(* IEC 61131-3 sources: RootPLC/demo/legacy-conveyor, 4 files *)

(* ---- 1-legacy.st ---- *)
PROGRAM PRG_Conveyor
VAR_INPUT start, stop, estop_ok : BOOL; speed_setpoint : INT; END_VAR
VAR_OUTPUT motor : BOOL; speed_cmd : SINT; jam_alarm : BOOL; END_VAR
VAR jam_timer : TON; jam_sensor : BOOL; END_VAR
motor := start OR motor AND NOT stop AND estop_ok;
speed_cmd := speed_setpoint;
jam_timer(IN := jam_sensor, PT := 3000);
IF jam_timer.Q THEN jam_alarm := 1; END_IF
END_PROGRAM

(* ---- 2-types-fixed.st ---- *)
(* The "obvious" fix: make the compiler happy, change nothing else. *)
PROGRAM PRG_Conveyor
VAR_INPUT start, stop, estop_ok, jam_sensor, reset : BOOL; speed_setpoint : INT; END_VAR
VAR_OUTPUT motor : BOOL; speed_cmd : SINT; jam_alarm : BOOL; END_VAR
VAR jam_timer : TON; END_VAR
motor := start OR motor AND NOT stop AND estop_ok;
speed_cmd := INT_TO_SINT(speed_setpoint);
jam_timer(IN := jam_sensor, PT := T#3s);
IF jam_timer.Q THEN jam_alarm := TRUE; END_IF
END_PROGRAM

(* ---- 3-correct.st ---- *)
PROGRAM PRG_Conveyor
VAR_INPUT
    start, stop, estop_ok, jam_sensor, reset : BOOL;
    speed_setpoint : INT;
END_VAR
VAR_OUTPUT
    motor, jam_alarm : BOOL;
    speed_cmd : SINT;
END_VAR
VAR
    jam_timer : TON;
END_VAR
jam_timer(IN := jam_sensor, PT := T#3s);
IF jam_timer.Q THEN
    jam_alarm := TRUE;
ELSIF reset THEN
    jam_alarm := FALSE;
END_IF
IF stop OR NOT estop_ok OR jam_alarm THEN
    motor := FALSE;
ELSIF start THEN
    motor := TRUE;
END_IF
IF motor THEN
    speed_cmd := INT_TO_SINT(LIMIT(0, speed_setpoint, 100));
ELSE
    speed_cmd := 0;
END_IF
END_PROGRAM

(* ---- safety_tests.st ---- *)
TEST safety_stop_wins_while_start_held
VAR uut : PRG_Conveyor; END_VAR
uut(start := TRUE, estop_ok := TRUE, speed_setpoint := 50);
uut(start := TRUE, stop := TRUE);
ASSERT_FALSE(uut.motor);
ASSERT_TRUE(uut.speed_cmd = 0);
END_TEST

TEST safety_estop_wins_and_needs_new_start
VAR uut : PRG_Conveyor; END_VAR
uut(start := TRUE, estop_ok := TRUE, speed_setpoint := 50);
uut(start := TRUE, estop_ok := FALSE);
ASSERT_FALSE(uut.motor);
uut(start := FALSE, estop_ok := TRUE);
ASSERT_FALSE(uut.motor);
uut(start := TRUE);
ASSERT_TRUE(uut.motor);
END_TEST

TEST safety_speed_is_clamped
VAR uut : PRG_Conveyor; END_VAR
uut(start := TRUE, estop_ok := TRUE, speed_setpoint := 250);
ASSERT_TRUE(uut.speed_cmd = 100);
uut(speed_setpoint := -40);
ASSERT_TRUE(uut.speed_cmd = 0);
uut(speed_setpoint := 75);
ASSERT_TRUE(uut.speed_cmd = 75);
END_TEST

TEST safety_jam_alarm_after_3s_latches
VAR uut : PRG_Conveyor; i : INT; END_VAR
uut(start := TRUE, estop_ok := TRUE, speed_setpoint := 50);
FOR i := 1 TO 25 DO
    uut(start := FALSE, jam_sensor := TRUE);
    ADVANCE(T#100ms);
END_FOR
ASSERT_FALSE(uut.jam_alarm);
ASSERT_TRUE(uut.motor);
FOR i := 1 TO 10 DO
    uut(jam_sensor := TRUE);
    ADVANCE(T#100ms);
END_FOR
uut(jam_sensor := FALSE);
ASSERT_TRUE(uut.jam_alarm);
ASSERT_FALSE(uut.motor);
uut(jam_sensor := FALSE);
ASSERT_TRUE(uut.jam_alarm);
uut(reset := TRUE);
ASSERT_FALSE(uut.jam_alarm);
END_TEST
